Fanuc KAREL source: kx00022.KL

-- PROVISIONAL review KL for V940-1; original PC SHA256 420fd8f4ca31b75c1c1371055fa3306997e6a6d4b75e3ff5d59439cc61f4ff7c
-- Incomplete behavior may be omitted. Consult companion uncertainty JSON. Do not deploy.
PROGRAM KX00022
%NOLOCKGROUP
VAR
  I : INTEGER
  J : INTEGER
  B : BOOLEAN
  F : FILE
  S : STRING[80]
-- UNRESOLVED_DECL P type=000102
-- UNRESOLVED_DECL BA type=002012
BEGIN
  -- V9_ZERO_TABLE_METADATA_HINT layout=0001; no indexed target words; source/name/runtime held
  -- UNRESOLVED_PC offsets 5-15; opcodes 9D,22,9D,33,35
  -- UNRESOLVED_PC offsets 20-35; opcodes 22,9D,33,34,23
  -- UNRESOLVED_PC offsets 40-44; opcodes 7F
END KX00022
